Omron CX-Programmer project NewProject (CX-Programmer 9.81)

# PLC NewPLC1: CJ2M CPU32
I/O table (CPU CJ2M-CPU32): rack 0 slot 11 CJ2M-EIP21

## Global symbols (name address type ; comment)
At_Entry 2.00 BOOL  ; At Entry
At_Exit 2.01 BOOL  ; At Exit
At_Load 2.02 BOOL  ; At Load
At_Unload 2.03 BOOL  ; At Unload
Emergency_stop 2.04 BOOL  ; Emergency stop
Entry_Conveyor 3.00 BOOL  ; Entry Conveyor
Exit_Conveyor 3.01 BOOL  ; Exit Conveyor
Load_Conveyor 3.02 BOOL  ; Load Conveyor
Reset 2.07 BOOL  ; Reset
Reset_light 3.06 BOOL  ; Reset light
Stacker_Crane_1_Left 3.08 BOOL  ; Stacker Crane 1 (Left)
Stacker_Crane_1_Left_Limit 2.10 BOOL  ; Stacker Crane 1 Left Limit
Stacker_Crane_1_Lift 3.07 BOOL  ; Stacker Crane 1 Lift
Stacker_Crane_1_Middle_Limit 2.12 BOOL  ; Stacker Crane 1 Middle Limit
Stacker_Crane_1_Moving_X 2.08 BOOL  ; Stacker Crane 1 Moving-X
Stacker_Crane_1_Moving_Z 2.09 BOOL  ; Stacker Crane 1 Moving-Z
Stacker_Crane_1_Right 3.09 BOOL  ; Stacker Crane 1 (Right)
Stacker_Crane_1_Right_Limit 2.11 BOOL  ; Stacker Crane 1 Right Limit
Stacker_Crane_1_Target_Pos_0 3.10 BOOL  ; Stacker Crane 1 Target Position Bool 0
Stacker_Crane_1_Target_Pos_1 3.11 BOOL  ; Stacker Crane 1 Target Position Bool 1
Stacker_Crane_1_Target_Pos_2 3.12 BOOL  ; Stacker Crane 1 Target Position Bool 2
Stacker_Crane_1_Target_Pos_3 3.13 BOOL  ; Stacker Crane 1 Target Position Bool 3
Stacker_Crane_1_Target_Pos_4 3.14 BOOL  ; Stacker Crane 1 Target Position Bool 4
Stacker_Crane_1_Target_Pos_5 3.15 BOOL  ; Stacker Crane 1 Target Position Bool 5
Start 2.05 BOOL  ; Start
Start_light 3.04 BOOL  ; Start light
Stop 2.06 BOOL  ; Stop
Stop_light 3.05 BOOL  ; Stop light
Unload_Conveyor 3.03 BOOL  ; Unload Conveyor
actual W0 UINT
enable W4.00 BOOL
i W200 UINT
load W4.01 BOOL
places W100 UINT[5]

## Program NewProgram1 (cyclic task 0)
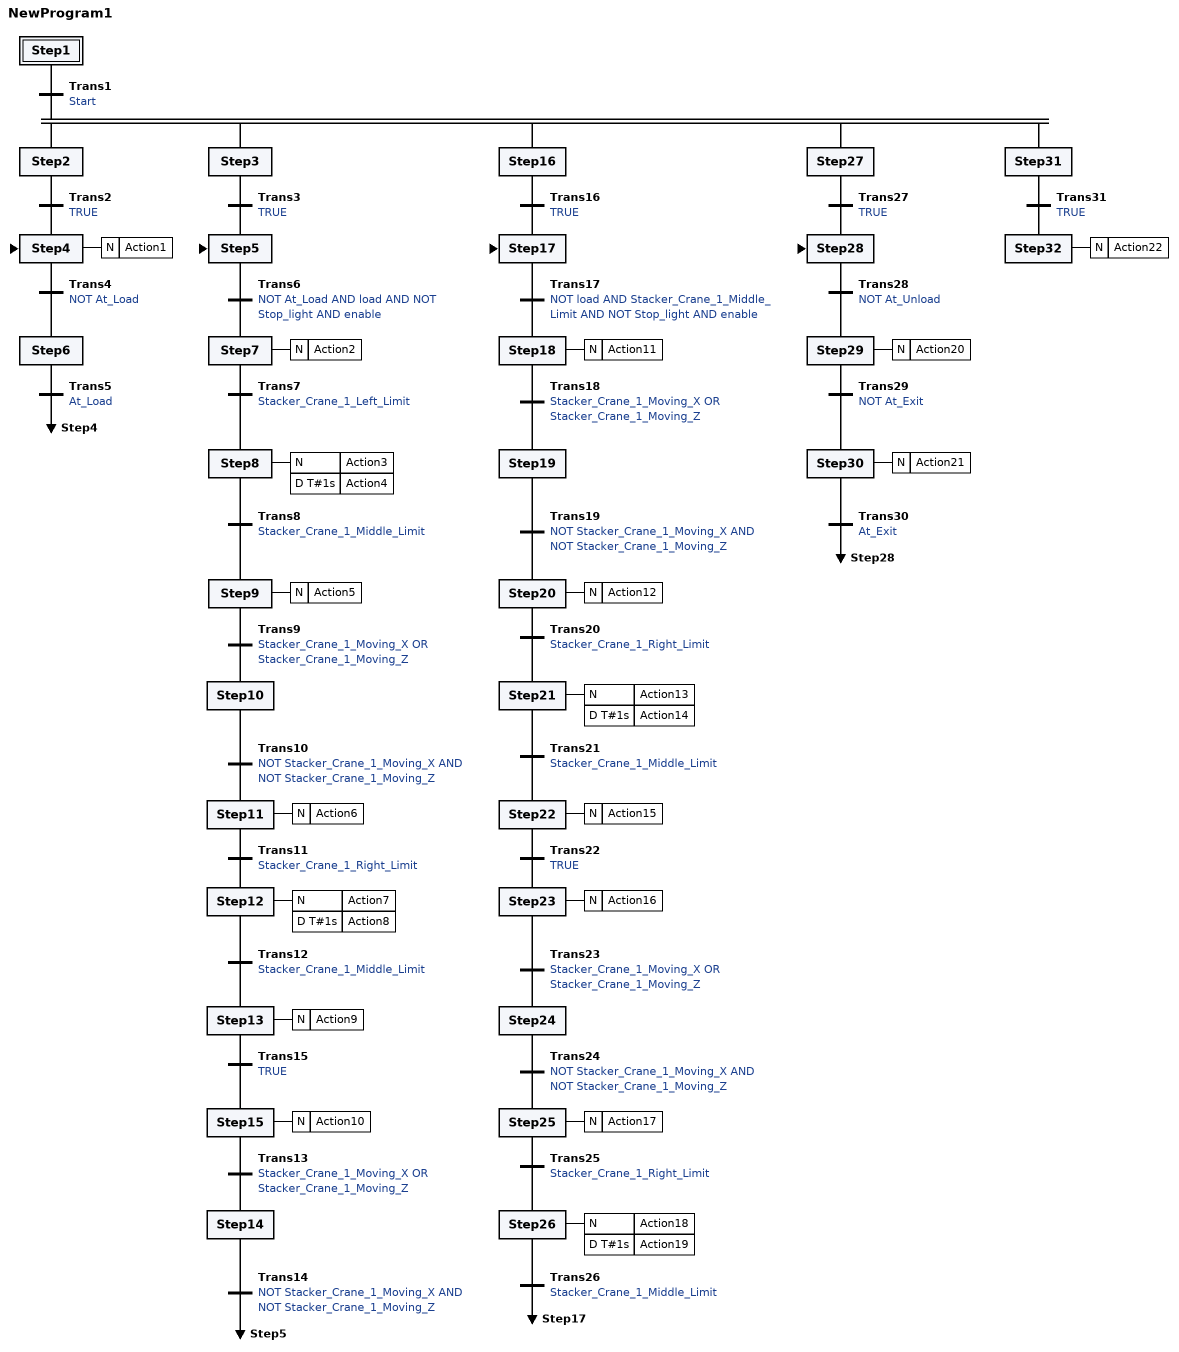
INITIAL_STEP Step1 :
END_STEP
TRANSITION Trans1 FROM Step1 TO (Step2,Step3,Step16,Step27,Step31)
 := Start;
END_TRANSITION
STEP Step2 :
END_STEP
STEP Step3 :
END_STEP
TRANSITION Trans2 FROM Step2 TO Step4
 := TRUE;
END_TRANSITION
STEP Step4 :
Action1(N) ;
END_STEP
TRANSITION Trans3 FROM Step3 TO Step5
 := TRUE;
END_TRANSITION
STEP Step5 :
END_STEP
TRANSITION Trans4 FROM Step4 TO Step6
 := NOT At_Load;
END_TRANSITION
STEP Step6 :
END_STEP
TRANSITION Trans5 FROM Step6 TO Step4
 := At_Load;
END_TRANSITION
TRANSITION Trans6 FROM Step5 TO Step7
 := NOT At_Load AND load AND NOT Stop_light AND enable;
END_TRANSITION
STEP Step7 :
Action2(N) ;
END_STEP
TRANSITION Trans7 FROM Step7 TO Step8
 := Stacker_Crane_1_Left_Limit;
END_TRANSITION
STEP Step8 :
Action3(N) ;
Action4(D,T#1s) ;
END_STEP
TRANSITION Trans8 FROM Step8 TO Step9
 := Stacker_Crane_1_Middle_Limit;
END_TRANSITION
STEP Step9 :
Action5(N) ;
END_STEP
TRANSITION Trans9 FROM Step9 TO Step10
 := Stacker_Crane_1_Moving_X OR Stacker_Crane_1_Moving_Z;
END_TRANSITION
STEP Step10 :
END_STEP
TRANSITION Trans10 FROM Step10 TO Step11
 := NOT Stacker_Crane_1_Moving_X AND NOT Stacker_Crane_1_Moving_Z;
END_TRANSITION
STEP Step11 :
Action6(N) ;
END_STEP
TRANSITION Trans11 FROM Step11 TO Step12
 := Stacker_Crane_1_Right_Limit;
END_TRANSITION
STEP Step12 :
Action7(N) ;
Action8(D,T#1s) ;
END_STEP
TRANSITION Trans12 FROM Step12 TO Step13
 := Stacker_Crane_1_Middle_Limit;
END_TRANSITION
STEP Step13 :
Action9(N) ;
END_STEP
TRANSITION Trans13 FROM Step15 TO Step14
 := Stacker_Crane_1_Moving_X OR Stacker_Crane_1_Moving_Z;
END_TRANSITION
STEP Step14 :
END_STEP
TRANSITION Trans14 FROM Step14 TO Step5
 := NOT Stacker_Crane_1_Moving_X AND NOT Stacker_Crane_1_Moving_Z;
END_TRANSITION
TRANSITION Trans15 FROM Step13 TO Step15
 := TRUE;
END_TRANSITION
STEP Step15 :
Action10(N) ;
END_STEP
STEP Step16 :
END_STEP
TRANSITION Trans16 FROM Step16 TO Step17
 := TRUE;
END_TRANSITION
STEP Step17 :
END_STEP
TRANSITION Trans17 FROM Step17 TO Step18
 := NOT load AND Stacker_Crane_1_Middle_Limit AND NOT Stop_light AND enable;
END_TRANSITION
STEP Step18 :
Action11(N) ;
END_STEP
TRANSITION Trans18 FROM Step18 TO Step19
 := Stacker_Crane_1_Moving_X OR Stacker_Crane_1_Moving_Z;
END_TRANSITION
STEP Step19 :
END_STEP
TRANSITION Trans19 FROM Step19 TO Step20
 := NOT Stacker_Crane_1_Moving_X AND NOT Stacker_Crane_1_Moving_Z;
END_TRANSITION
STEP Step20 :
Action12(N) ;
END_STEP
TRANSITION Trans20 FROM Step20 TO Step21
 := Stacker_Crane_1_Right_Limit;
END_TRANSITION
STEP Step21 :
Action13(N) ;
Action14(D,T#1s) ;
END_STEP
TRANSITION Trans21 FROM Step21 TO Step22
 := Stacker_Crane_1_Middle_Limit;
END_TRANSITION
STEP Step22 :
Action15(N) ;
END_STEP
TRANSITION Trans22 FROM Step22 TO Step23
 := TRUE;
END_TRANSITION
STEP Step23 :
Action16(N) ;
END_STEP
TRANSITION Trans23 FROM Step23 TO Step24
 := Stacker_Crane_1_Moving_X OR Stacker_Crane_1_Moving_Z;
END_TRANSITION
STEP Step24 :
END_STEP
TRANSITION Trans24 FROM Step24 TO Step25
 := NOT Stacker_Crane_1_Moving_X AND NOT Stacker_Crane_1_Moving_Z;
END_TRANSITION
STEP Step25 :
Action17(N) ;
END_STEP
TRANSITION Trans25 FROM Step25 TO Step26
 := Stacker_Crane_1_Right_Limit;
END_TRANSITION
STEP Step26 :
Action18(N) ;
Action19(D,T#1s) ;
END_STEP
TRANSITION Trans26 FROM Step26 TO Step17
 := Stacker_Crane_1_Middle_Limit;
END_TRANSITION
STEP Step27 :
END_STEP
TRANSITION Trans27 FROM Step27 TO Step28
 := TRUE;
END_TRANSITION
STEP Step28 :
END_STEP
TRANSITION Trans28 FROM Step28 TO Step29
 := NOT At_Unload;
END_TRANSITION
STEP Step29 :
Action20(N) ;
END_STEP
TRANSITION Trans29 FROM Step29 TO Step30
 := NOT At_Exit;
END_TRANSITION
STEP Step30 :
Action21(N) ;
END_STEP
TRANSITION Trans30 FROM Step30 TO Step28
 := At_Exit;
END_TRANSITION
STEP Step31 :
END_STEP
TRANSITION Trans31 FROM Step31 TO Step32
 := TRUE;
END_TRANSITION
STEP Step32 :
Action22(N) ;
END_STEP

### Action Action1

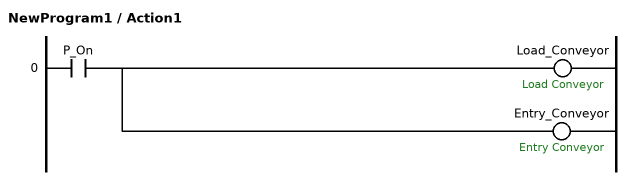
; rung 0
LD P_On
OUT Load_Conveyor  ; Load Conveyor
OUT Entry_Conveyor  ; Entry Conveyor

### Action Action2

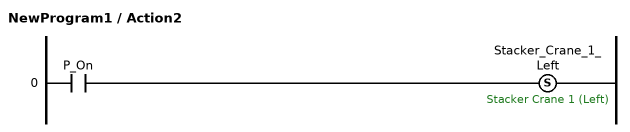
; rung 0
LD P_On
SET Stacker_Crane_1_Left  ; Stacker Crane 1 (Left)

### Action Action3

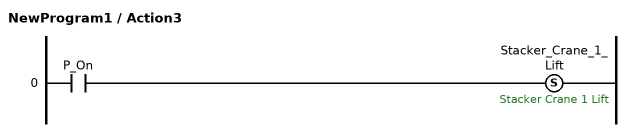
; rung 0
LD P_On
SET Stacker_Crane_1_Lift  ; Stacker Crane 1 Lift

### Action Action4

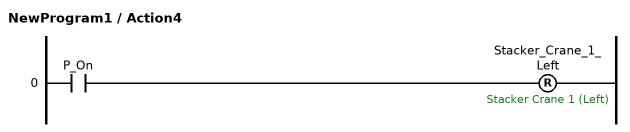
; rung 0
LD P_On
RSET Stacker_Crane_1_Left  ; Stacker Crane 1 (Left)

### Action Action5

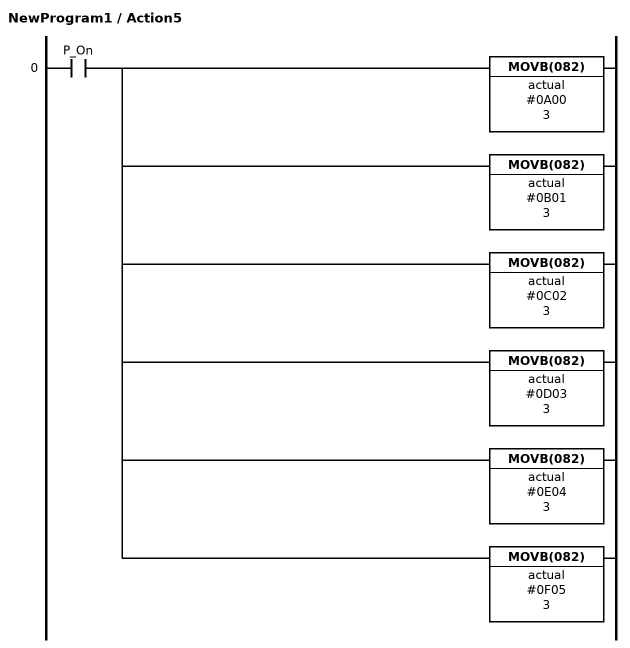
; rung 0
LD P_On
MOVB(082) actual #0A00 3
MOVB(082) actual #0B01 3
MOVB(082) actual #0C02 3
MOVB(082) actual #0D03 3
MOVB(082) actual #0E04 3
MOVB(082) actual #0F05 3

### Action Action6

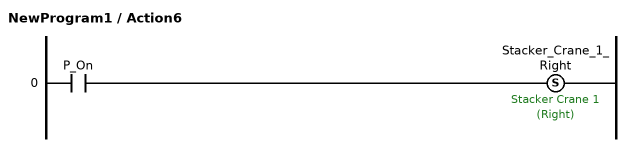
; rung 0
LD P_On
SET Stacker_Crane_1_Right  ; Stacker Crane 1 (Right)

### Action Action7

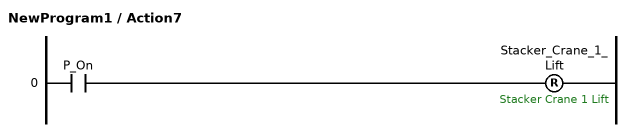
; rung 0
LD P_On
RSET Stacker_Crane_1_Lift  ; Stacker Crane 1 Lift

### Action Action8

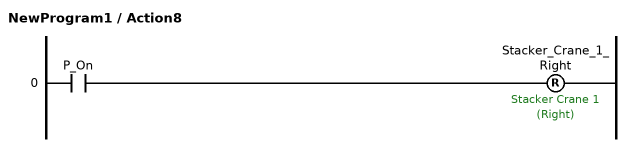
; rung 0
LD P_On
RSET Stacker_Crane_1_Right  ; Stacker Crane 1 (Right)

### Action Action9

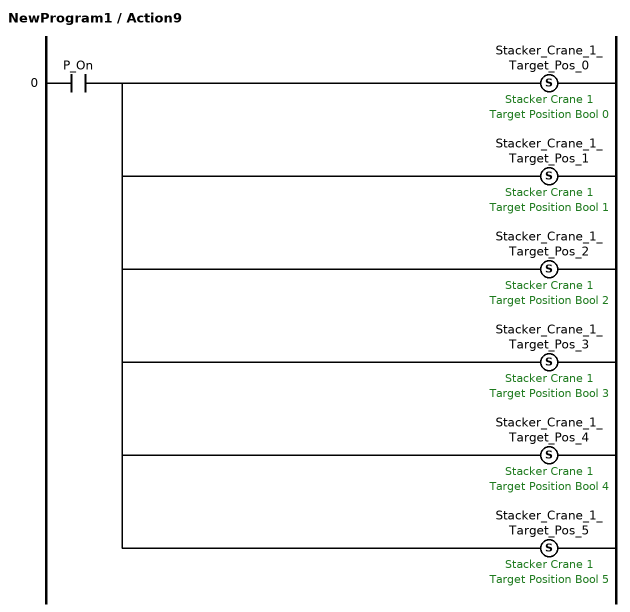
; rung 0
LD P_On
SET Stacker_Crane_1_Target_Pos_0  ; Stacker Crane 1 Target Position Bool 0
SET Stacker_Crane_1_Target_Pos_1  ; Stacker Crane 1 Target Position Bool 1
SET Stacker_Crane_1_Target_Pos_2  ; Stacker Crane 1 Target Position Bool 2
SET Stacker_Crane_1_Target_Pos_3  ; Stacker Crane 1 Target Position Bool 3
SET Stacker_Crane_1_Target_Pos_4  ; Stacker Crane 1 Target Position Bool 4
SET Stacker_Crane_1_Target_Pos_5  ; Stacker Crane 1 Target Position Bool 5

### Action Action10

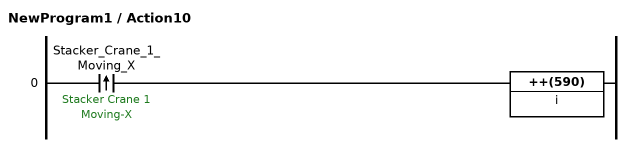
; rung 0
@LD Stacker_Crane_1_Moving_X  ; Stacker Crane 1 Moving-X
++(590) i

### Action Action11

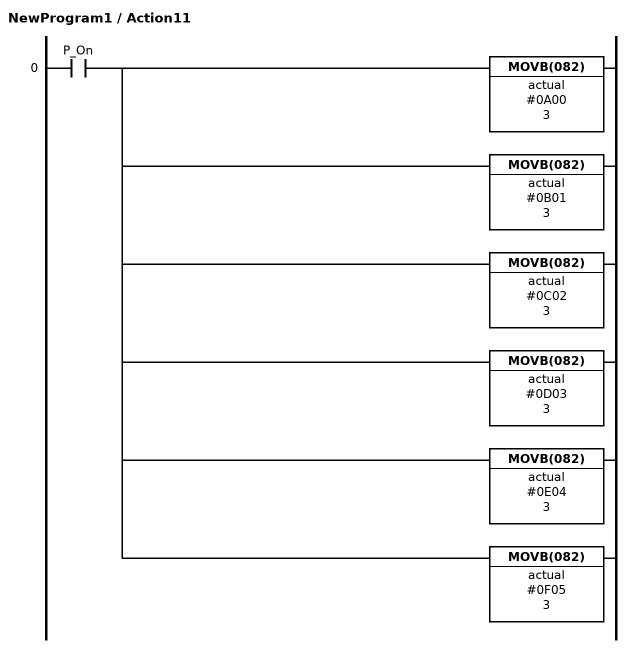
; rung 0
LD P_On
MOVB(082) actual #0A00 3
MOVB(082) actual #0B01 3
MOVB(082) actual #0C02 3
MOVB(082) actual #0D03 3
MOVB(082) actual #0E04 3
MOVB(082) actual #0F05 3

### Action Action12

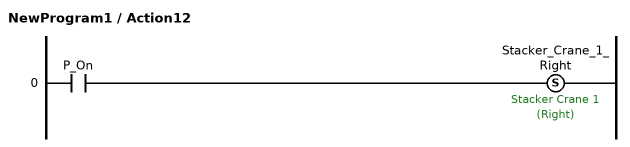
; rung 0
LD P_On
SET Stacker_Crane_1_Right  ; Stacker Crane 1 (Right)

### Action Action13

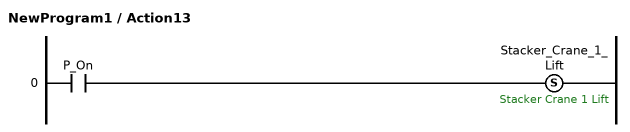
; rung 0
LD P_On
SET Stacker_Crane_1_Lift  ; Stacker Crane 1 Lift

### Action Action14

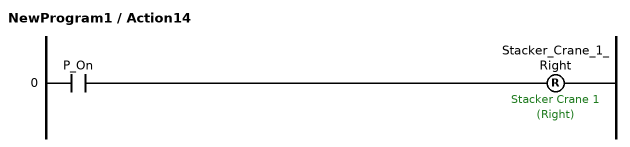
; rung 0
LD P_On
RSET Stacker_Crane_1_Right  ; Stacker Crane 1 (Right)

### Action Action15

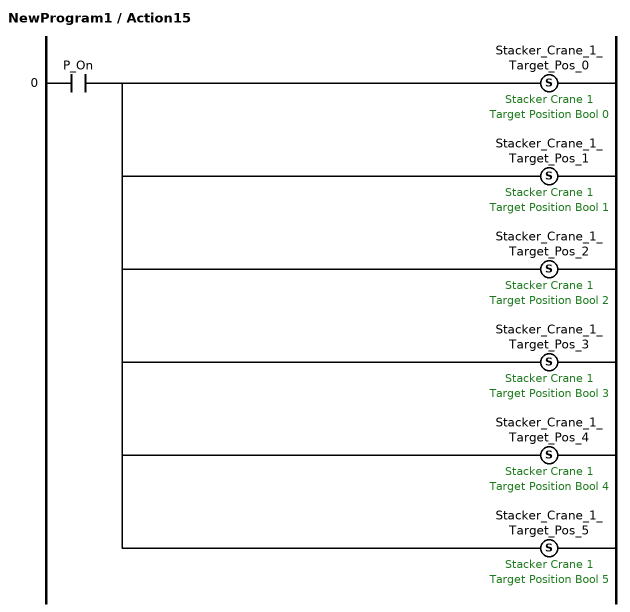
; rung 0
LD P_On
SET Stacker_Crane_1_Target_Pos_0  ; Stacker Crane 1 Target Position Bool 0
SET Stacker_Crane_1_Target_Pos_1  ; Stacker Crane 1 Target Position Bool 1
SET Stacker_Crane_1_Target_Pos_2  ; Stacker Crane 1 Target Position Bool 2
SET Stacker_Crane_1_Target_Pos_3  ; Stacker Crane 1 Target Position Bool 3
SET Stacker_Crane_1_Target_Pos_4  ; Stacker Crane 1 Target Position Bool 4
SET Stacker_Crane_1_Target_Pos_5  ; Stacker Crane 1 Target Position Bool 5

### Action Action16

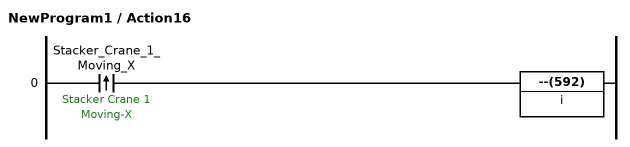
; rung 0
@LD Stacker_Crane_1_Moving_X  ; Stacker Crane 1 Moving-X
--(592) i

### Action Action17

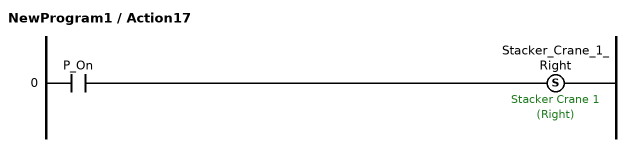
; rung 0
LD P_On
SET Stacker_Crane_1_Right  ; Stacker Crane 1 (Right)

### Action Action18

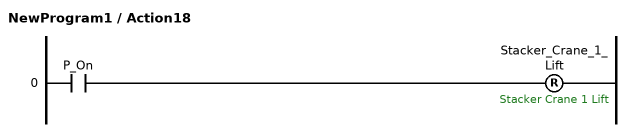
; rung 0
LD P_On
RSET Stacker_Crane_1_Lift  ; Stacker Crane 1 Lift

### Action Action19

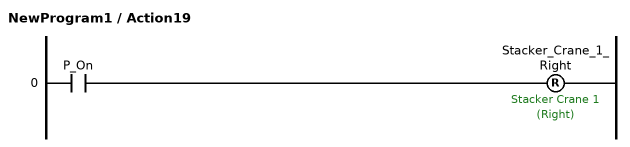
; rung 0
LD P_On
RSET Stacker_Crane_1_Right  ; Stacker Crane 1 (Right)

### Action Action20

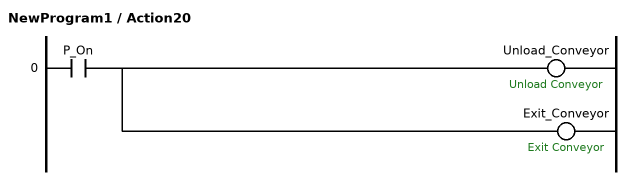
; rung 0
LD P_On
OUT Unload_Conveyor  ; Unload Conveyor
OUT Exit_Conveyor  ; Exit Conveyor

### Action Action21

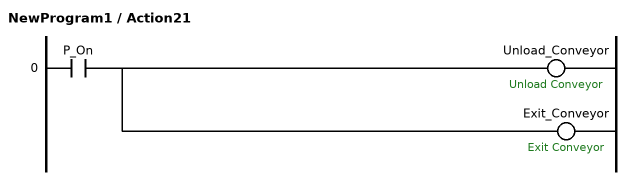
; rung 0
LD P_On
OUT Unload_Conveyor  ; Unload Conveyor
OUT Exit_Conveyor  ; Exit Conveyor

### Action Action22

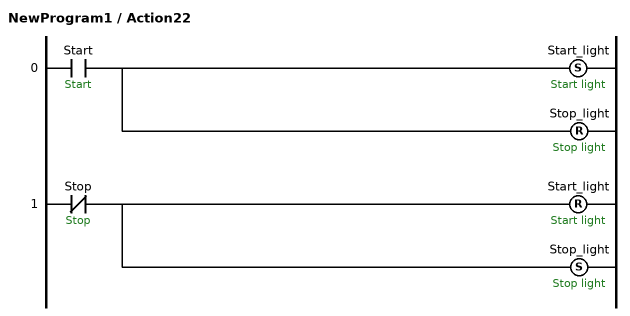
; rung 0
LD Start  ; Start
SET Start_light  ; Start light
RSET Stop_light  ; Stop light
; rung 1
LDNOT Stop  ; Stop
RSET Start_light  ; Start light
SET Stop_light  ; Stop light

## Program NewProgram2 (cyclic task 1)
IF P_First_Cycle THEN
	i:=0;
	places[0] := 1;
	places[1] := 7;
	places[2] := 19;
	places[3] := 30;
	places[4] := 50;
	
	actual := 0;
	load := TRUE;
	enable :=  TRUE;
END_IF;

actual := places[i];

IF i = 5 THEN
	load := FALSE;
	i := i-1;
END_IF;


IF NOT load AND i>5 THEN
	enable:= FALSE;
END_IF;